Fanuc KAREL source: KO00039.KL

PROGRAM KO00039
%NOLOCKGROUP
%ENVIRONMENT MIR
VAR
  P1: POSITION
  P2: XYZWPR
  F: BOOLEAN
  OUT: XYZWPREXT
BEGIN
  F = TRUE
  OUT = MIRROR(P1, P2, F)
END KO00039
